          MoveL speed 75 mm/s, acceleration 150 mm/s^2 (useActiveTCP=true) feature=FRM_Reference
            SuppressedNode
              Script: PSE_T[2]=PSE_T[2]-0.005
            Waypoint Variable (Variable): variable=PSE_T
            SuppressedNode
              Force Frame feature=FRM_Reference; selection=[1, 1, 0, 0, 0, 0]; wrench=[0, 0, 0, 0, 0, 0]; limitsForce=[0.25, 0.25, 0.15, 1.047198, 1.047198, 1.047198]; limitsMotion=[0.1, 0.1, 0.1, 0.349066, 0.349066, 0.349066]
                Waypoint Variable (Variable): motionParameters(jointSpeed=1.047198 jointAcceleration=1.396263 cartesianSpeed=0.03 cartesianAcceleration=0.2); variable=PSE_T
            'ADD OPEN GRIPPER'
            Script: rq_set_force_norm(20)
            Script: rq_set_speed_norm(30)
            Script: rq_move_and_wait_norm(GRP_Close_Pos)
          Set DigitalOutput pin=digital_out[4]; digitalValue=1
          Wait Sleep waitTime=0.3
          MoveL speed 100 mm/s, acceleration 1200 mm/s^2 (useActiveTCP=true) feature=FRM_Reference
            Waypoint Variable (Variable): motionParameters(jointSpeed=1.047198 jointAcceleration=1.396263 cartesianSpeed=0.25 cartesianAcceleration=1.2); variable=PSE_R
      Case (caseValue=4)
        Folder Place probe in 3finger
          Action_Info := "place object"
          MoveJ speed 100 deg/s, acceleration 80 deg/s^2 (useActiveTCP=true) feature=FRM_Reference
            Waypoint Variable (Variable): variable=PSE_A
          Set DigitalOutput pin=digital_out[4]; digitalValue=1
          MoveL speed 75 mm/s, acceleration 150 mm/s^2 (useActiveTCP=true) feature=FRM_Reference
            Waypoint Variable (Variable): variable=PSE_T
              Until TOOL_CONTACT_DETECTION (allowActions=false retraction=0 decelerationAcceleration=3 decelerationAngularAcceleration=34.906585)
          Set DigitalOutput pin=digital_out[4]; digitalValue=0
          Wait Sleep waitTime=0.5
          SuppressedNode
            If Task_ID≟12
              Wait Sleep waitTime=0.15
              MoveL speed 75 mm/s, acceleration 150 mm/s^2 (useActiveTCP=true) feature=FRM_Reference
                Waypoint Variable (Variable): variable=PSE_R
      Case (caseValue=5)
        SuppressedNode
          Folder Decapping
            Action_Info := "decapping"
            PRM_decap_Zval := z_Pos
            PRM_forcdistSta := 0.02
            Script: zero_ftsensor()
            Wait Sleep waitTime=1
            Set DigitalOutput pin=digital_out[5]; digitalValue=1
            Set DigitalOutput pin=digital_out[3]; digitalValue=1
            Force Frame feature=uML_3fingergrip; selection=[0, 0, 1, 0, 0, 0]; wrench=[0, 0, 5, 0, 0, 0]; limitsForce=[0.04, 0.04, 0.015, 1.047198, 1.047198, 1.047198]; limitsMotion=[0.1, 0.1, 0.1, 0.349066, 0.349066, 0.349066]
              PRC_Force_Decap := True
              Wait Condition expression=PRM_forcdistLiv>PRM_forcdistSta
            PRC_Force_Decap := False
            Set DigitalOutput pin=digital_out[5]; digitalValue=0
            Set DigitalOutput pin=digital_out[3]; digitalValue=0
            MoveL speed 150 mm/s, acceleration 800 mm/s^2 (useActiveTCP=true) feature=FRM_Reference
              Waypoint Variable (Variable): variable=PSE_R
        Folder Decapping
          Action_Info := "decapping"
          Set DigitalOutput pin=digital_out[5]; digitalValue=1
          Set DigitalOutput pin=digital_out[3]; digitalValue=1
          Script: action_manipulator_decapping()
          Set DigitalOutput pin=digital_out[5]; digitalValue=0
          Set DigitalOutput pin=digital_out[3]; digitalValue=0
          MoveL speed 150 mm/s, acceleration 800 mm/s^2 (useActiveTCP=true) feature=FRM_Reference
            Waypoint Variable (Variable): variable=PSE_R
      Case (caseValue=6)
        SuppressedNode
          Folder Drop the cap
            Script: rq_set_speed_norm(100)
            Script: rq_set_force_norm(10)
            MoveJ speed 100 deg/s, acceleration 80 deg/s^2 (useActiveTCP=true) feature=FRM_Reference
              Waypoint Variable (Variable): motionParameters(blendRadius=0.02); variable=PSE_A
            MoveL speed 400 mm/s, acceleration 500 mm/s^2 (useActiveTCP=true) feature=FRM_Reference
              Waypoint Variable (Variable): motionParameters(jointSpeed=1.047198 jointAcceleration=1.396263 cartesianSpeed=0.09 cartesianAcceleration=0.05); variable=PSE_T
              'ADD OPEN GRIPPER'
              Loop While (checkContinuously=false) expression=rq_is_object_detected()
                URCap Gripper (Robotiq_Grippers, Robotiq Inc.) dataModel(position=0.0, force=28.0, speed=100.0, positionInDouble=0.0, forceInDouble=28.0, speedInDouble=100.0, slaveIds=[9], blocking=true)
                Wait Sleep waitTime=0.01
                URCap Gripper (Robotiq_Grippers, Robotiq Inc.) dataModel(position=100.0, force=28.0, speed=100.0, positionInDouble=100.0, forceInDouble=28.0, speedInDouble=100.0, slaveIds=[9], blocking=true)
              Wait Sleep waitTime=0.2
              Waypoint Variable (Variable): variable=PSE_R
        Folder Drop
          Script: rq_set_speed_norm(100)
          MoveJ speed 100 deg/s, acceleration 80 deg/s^2 (useActiveTCP=true) feature=FRM_Reference
            Waypoint Variable (Variable): motionParameters(blendRadius=0.02); variable=PSE_A
          MoveL speed 400 mm/s, acceleration 500 mm/s^2 (useActiveTCP=true) feature=FRM_Reference
            Waypoint Variable (Variable): motionParameters(jointSpeed=1.047198 jointAcceleration=1.396263 cartesianSpeed=0.12 cartesianAcceleration=0.08); variable=PSE_T
            URCap Gripper (Robotiq_Grippers, Robotiq Inc.) dataModel(position=70.19607843137254, force=30.19607843137255, speed=0.0, positionInDouble=70.19607843137254, forceInDouble=30.19607843137255, speedInDouble=0.0, slaveIds=[9], blocking=true)
            Waypoint Variable (Variable): motionParameters(jointSpeed=1.047198 jointAcceleration=1.396263 cartesianSpeed=0.12 cartesianAcceleration=0.08); variable=PSE_T_H
            Script: rq_move_and_wait_norm(GRP_Open_Pos)
            Wait Sleep waitTime=0.2
            Waypoint Variable (Variable): variable=PSE_R
      Case (caseValue=7)
        Folder Load
          Action_Info := "load object in the machine"
          SuppressedNode
            Script: do_transition(keep_rxry=OBJ_Picked)
          If JNT_Q≠JNT_Z
            Script: movej(get_inverse_kin(pose_trans(FRM_Reference, PSE_A), qnear=JNT_Q), r=0.05)
          Else 
            MoveJ speed 100 deg/s, acceleration 80 deg/s^2 (useActiveTCP=true) feature=FRM_Reference
              Waypoint Variable (Variable): motionParameters(blendRadius=0.02); variable=PSE_A
          MoveL speed 400 mm/s, acceleration 500 mm/s^2 (useActiveTCP=true) feature=FRM_Reference
            SuppressedNode
              Waypoint Variable (Variable): motionParameters(jointSpeed=1.047198 jointAcceleration=1.396263 cartesianSpeed=0.09 cartesianAcceleration=0.05); variable=PSE_T
                Until TOOL_CONTACT_DETECTION (allowActions=false retraction=0 decelerationAcceleration=0.5 decelerationAngularAcceleration=34.906585)
            SuppressedNode
              Force Frame feature=FRM_Reference; selection=[1, 1, 0, 0, 0, 0]; wrench=[0, 0, 0, 0, 0, 0]; limitsForce=[0.05, 0.05, 0.15, 1.047198, 1.047198, 1.047198]; limitsMotion=[0.1, 0.1, 0.1, 0.349066, 0.349066, 0.349066]
                Waypoint Variable (Variable): motionParameters(jointSpeed=1.047198 jointAcceleration=1.396263 cartesianSpeed=0.07 cartesianAcceleration=0.04); variable=PSE_T
            Waypoint Variable (Variable): motionParameters(jointSpeed=1.047198 jointAcceleration=1.396263 cartesianSpeed=0.07 cartesianAcceleration=0.04); variable=PSE_T_H
            URCap Gripper (Robotiq_Grippers, Robotiq Inc.) dataModel(position=100.0, force=0.0, speed=67.84313725490196, positionInDouble=100.0, forceInDouble=0.0, speedInDouble=67.84313725490196, slaveIds=[9], blocking=true)
            Wait Sleep waitTime=0.2
            Waypoint Variable (Variable): motionParameters(jointSpeed=1.047198 jointAcceleration=1.396263 cartesianSpeed=0.07 cartesianAcceleration=0.04); variable=PSE_T
            Waypoint Variable (Variable): variable=PSE_R
      Case (caseValue=8)
        Folder UnLoad
          Action_Info := "unload object in the machine"
          SuppressedNode
            Script: do_transition(keep_rxry=OBJ_Picked)
          If JNT_Q≠JNT_Z
            SuppressedNode
              Script: movej(get_inverse_kin(pose_trans(FRM_Reference, PSE_A), qnear=JNT_Q), r=0.01)
            Script: movej(get_inverse_kin(pose_trans(FRM_Reference, PSE_A), qnear=JNT_Q))
          Else 
            MoveJ speed 100 deg/s, acceleration 80 deg/s^2 (useActiveTCP=true) feature=FRM_Reference
              Waypoint Variable (Variable): variable=PSE_A
          MoveL speed 400 mm/s, acceleration 500 mm/s^2 (useActiveTCP=true) feature=FRM_Reference
            SuppressedNode
              Waypoint Variable (Variable): motionParameters(jointSpeed=1.047198 jointAcceleration=1.396263 cartesianSpeed=0.09 cartesianAcceleration=0.05); variable=PSE_T
                Until TOOL_CONTACT_DETECTION (allowActions=false retraction=0 decelerationAcceleration=0.5 decelerationAngularAcceleration=34.906585)
            SuppressedNode
              Force Frame feature=FRM_Reference; selection=[1, 1, 0, 0, 0, 0]; wrench=[0, 0, 0, 0, 0, 0]; limitsForce=[0.05, 0.05, 0.15, 1.047198, 1.047198, 1.047198]; limitsMotion=[0.1, 0.1, 0.1, 0.349066, 0.349066, 0.349066]
                Waypoint Variable (Variable): motionParameters(jointSpeed=1.047198 jointAcceleration=1.396263 cartesianSpeed=0.07 cartesianAcceleration=0.04); variable=PSE_T
            Script: rq_move_and_wait_norm(GRP_Open_Pos)
            Waypoint Variable (Variable): motionParameters(jointSpeed=1.047198 jointAcceleration=1.396263 cartesianSpeed=0.07 cartesianAcceleration=0.04); variable=PSE_T_H
            URCap Gripper (Robotiq_Grippers, Robotiq Inc.) dataModel(position=100.0, force=0.0, speed=67.84313725490196, positionInDouble=100.0, forceInDouble=0.0, speedInDouble=67.84313725490196, slaveIds=[9], blocking=true)
            Wait Sleep waitTime=0.2
            OBJ_Picked := rq_is_object_detected()
            If OBJ_Picked
              Waypoint Variable (Variable): motionParameters(jointSpeed=1.047198 jointAcceleration=1.396263 cartesianSpeed=0.07 cartesianAcceleration=0.04); variable=PSE_T
              Script: rq_move_and_wait_norm(GRP_Open_Pos)
              Waypoint Variable (Variable): variable=PSE_R
            Else 
              Script: set_error(1010)
      Case (caseValue=16)
        Folder Scan the barcode
          Action_Info := "scan the barcode"
          Barc_scan_succs := False
          Folder First check
            Set DigitalOutput pin=digital_out[6]; digitalValue=1
            Wait Sleep waitTime=0.1
            Barc_scan_succs := digital_in[6]
          If Barc_scan_succs
            Set DigitalOutput pin=digital_out[5]; digitalValue=1
            Set DigitalOutput pin=digital_out[2]; digitalValue=1
            Loop While (checkContinuously=true) expression=Barc_scan_succs
              Barc_scan_succs := digital_in[6]
              Wait Sleep waitTime=0.05
            Set DigitalOutput pin=digital_out[5]; digitalValue=0
            Set DigitalOutput pin=digital_out[2]; digitalValue=0
            Set DigitalOutput pin=digital_out[6]; digitalValue=0
          Else 
            Timer (action=Reset) variable=Timer_Barc_scan
            Timer (action=Start) variable=Timer_Barc_scan
            Set DigitalOutput pin=digital_out[3]; digitalValue=1
            Set DigitalOutput pin=digital_out[5]; digitalValue=1
            Loop While (checkContinuously=true) expression=not Barc_scan_succs and  not CMD_Stop and Timer_Barc_scan<60
              SuppressedNode
                If Timer_Barc_scan>1.5
                  Placeholder
              Set DigitalOutput pin=digital_out[6]; digitalValue=1
              Barc_scan_succs := digital_in[6]
              Wait Sleep waitTime=0.05
            Set DigitalOutput pin=digital_out[5]; digitalValue=0
            Set DigitalOutput pin=digital_out[3]; digitalValue=0
            Set DigitalOutput pin=digital_out[6]; digitalValue=0
            Timer (action=Stop) variable=Timer_Barc_scan
            If Timer_Barc_scan≥60
              Script: set_error(5200)
    '=========='
    Script: textmsg("Action=",Action)
    Folder PostSettings [hidden by the author, left out]
SubProgram Sub_AMR_MiR_V3 [hidden by the author, left out]
SubProgram Sub_Action_V4 (keepSynchronizedWithDisk=true) programFile=/programs/03 Sub Routines/Sub_Action_V4.urp
  Folder PreSettings
    Folder init poses [hidden by the author, left out]
    Folder Gripping parameters
      Script: OBJ = find_object_by_type(OBJs, OBJ_Type)
      GRP_Open_Pos := OBJ.dimension.diameter * 1000 + 6
      GRP_Offset := OBJ.gripper_offset
      Script: rq_set_force_norm(50)
      Script: rq_set_speed_norm(50)
    Switch expression=ITM_ID
      Case (caseValue=1)
        Folder uML
          Script: JIG2 = find_object_by_type(JIGs, JIG)
          JIG_Offset := JIG2.jig_offset
          Switch expression=JIG
            Case (caseValue=1)
              Folder 3FG
                Folder define poses
                  FRM_Reference := ULM_3FG
                  JNT_Q := JNT_HOME
                  PSE_T := pose_trans(GRP_Offset, JIG_Offset)
                  PSE_A := pose_trans(PSE_T, p[0,0,0.100,0,0,0])
                  PSE_R := pose_add(PSE_T, p[0,0,0.100,0,0,0])
            Case (caseValue=2)
              Folder Input
                'CHANGE THE REFERENCE TO THE FRAME TO MOVE IN'
                Folder define poses
                  FRM_Reference := ULM_Input
                  PSE_T := pose_trans(pose_trans(get_pattern_pos_rectangle(OBJ_Nbr, "X", [10,5], patternsize=[0.181,0.081]), GRP_Offset), JIG_Offset)
                  If Action≟1
                    PSE_R := pose_add(PSE_T, p[0,0,0.200,0,0,0])
                    PSE_A := pose_add(PSE_T, p[0,0,0.100,0,0,0])
                  ElseIf Action≟2
                    PSE_R := pose_add(PSE_T, p[0,0,0.100,0,0,0])
                    PSE_A := pose_add(PSE_T, p[0,0,0.200,0,0,0])
            Case (caseValue=3)
              Folder Output
                'CHANGE THE REFERENCE TO THE FRAME TO MOVE IN'
                Folder define poses
                  FRM_Reference := ULM_Output
                  PSE_T := pose_trans(pose_trans(get_pattern_pos_rectangle(OBJ_Nbr, "X", [10,5], patternsize=[0.181,0.081]), GRP_Offset), JIG_Offset)
                  SuppressedNode
                    PSE_T_H := 
                  If Action≟1
                    PSE_R := pose_add(PSE_T, p[0,0,0.200,0,0,0])
                    PSE_A := pose_add(PSE_T, p[0,0,0.100,0,0,0])
                  ElseIf Action≟2
                    PSE_R := pose_add(PSE_T, p[0,0,0.100,0,0,0])
                    PSE_A := pose_add(PSE_T, p[0,0,0.200,0,0,0])
            Case (caseValue=4)
              Folder jig centrifuge racks
                Folder define poses
                  FRM_Reference := ULM_Cent_Racks
                  PSE_T := get_pattern_pos_rectangle(JIG_Slot, "X", [4,1], patternsize=[0.291,0])
                  If OBJ_Nbr≠0
                    PSE_T := pose_trans(pose_trans(PSE_T, get_pattern_pos_rectangle(OBJ_Nbr, "X", [3,3], patternsize=[0.060,0.060])),p[-0.030, -0.030,0,0,0,3.927])
                  PSE_T := pose_trans(PSE_T, GRP_Offset)
                  If Action≟1
                    PSE_R := pose_add(PSE_T, p[0,0,0.200,0,0,0])
                    PSE_A := pose_add(PSE_T, p[0,0,0.100,0,0,0])
                  ElseIf Action≟2
                    PSE_R := pose_add(PSE_T, p[0,0,0.100,0,0,0])
                    PSE_A := pose_add(PSE_T, p[0,0,0.200,0,0,0])
            Case (caseValue=6)
              Folder Caps bin
                Folder define poses
                  'Drop cap'
                  Script: FRM_Reference=ULM_Cap_Bin
                  PSE_T := pose_RPY2RotVec(p[0,0,0,0,0,0])
                  PSE_T_H := pose_add(PSE_T, p[0,0,-0.011,0,0,0])
                  PSE_A := pose_trans(PSE_T, p[0,0,0.1,0,0,0])
                  PSE_R := pose_add(PSE_T, p[0,0,0.100,0,0,0])
            Case (caseValue=7)
              Folder Sarstedt
                'CHANGE THE REFERENCE TO THE FRAME TO MOVE IN'
                SuppressedNode
                  Folder Gripping parameters
                    GRP_Open_Pos := 45
                    GRP_Close_Pos := 100
                    Script: rq_set_force_norm(80)
                    Script: rq_set_speed_norm(100)
                If TASK.ID≟10
                  Folder Frame & Position Params
                    Script: FRM_Reference = ULM_SS_Rack
                    SuppressedNode
                      MoveL speed 250 mm/s, acceleration 1200 mm/s^2 (useActiveTCP=true) feature=FRM_Reference
                        Waypoint Variable (Variable): variable(featureName=uLM_SS_PickPlc)
                    SuppressedNode
                      PSE_T := pose_RPY2RotVec(p[0,0,0,0,0,0])
                    SuppressedNode
                      PSE_T := pose_trans(PSE_T, GRP_Offset)
                    PSE_T := uLM_SS_PickPlc
                    PSE_A := pose_trans(PSE_T, p[0,0,0.1,0,0,0])
                    PSE_R := pose_add(PSE_T, p[0,0,0.1,0,0,0])
                ElseIf TASK.ID≟11
                  Script: FRM_Reference = uLM_SS_PickPlc
                  PSE_T := pose_RPY2RotVec(p[0,0,0,0,0,0])
                  PSE_T := pose_trans(PSE_T, GRP_Offset)
                  PSE_A := pose_trans(PSE_T, p[0,0,0.1,0,0,0])
                  PSE_R := pose_add(PSE_T, p[0,0,0.2,0,0,0])
      Case (caseValue=2)
        Folder Centrifuge
          'CHANGE THE REFERENCE TO THE FRAME TO MOVE IN'
          Folder define poses
            FRM_Reference := FRM_Centrifuge
            PSE_T := GRP_Offset
            If Action≟8
              PSE_R := pose_add(PSE_T, p[0,0,0.250,0,0,0])
              PSE_A := pose_add(PSE_T, p[0,0,0.150,0,0,0])
            ElseIf Action≟7
              PSE_R := pose_add(PSE_T, p[0,0,0.150,0,0,0])
              PSE_A := pose_add(PSE_T, p[0,0,0.250,0,0,0])
      Case (caseValue=3)
        Folder Output
          'CHANGE THE REFERENCE TO THE FRAME TO MOVE IN'
          Folder define poses
            FRM_Reference := Base
            PSE_T := p[0,0,0,0,0,0]
            PSE_A := pose_add(PSE_T, p[0,0,0.150,0,0,0])
            PSE_R := pose_add(PSE_T, p[0,0,0.100,0,0,0])
      Case (caseValue=5)
        Folder Sarstedt Pickup Table
          'CHANGE THE REFERENCE TO THE FRAME TO MOVE IN'
          Switch expression=JIG
            Case (caseValue=7)
              Folder Sarstedt Rack
                SuppressedNode
                  Folder Gripping parameters
                    GRP_Open_Pos := 45
                    GRP_Close_Pos := 100
                    Script: rq_set_force_norm(80)
                    Script: rq_set_speed_norm(100)
                Folder Frame & Position Params
                  Script: FRM_Reference = FRM_SS_SSTable
                  PSE_T := pose_RPY2RotVec(p[0,0,0,0,0,0])
                  PSE_T := pose_trans(PSE_T, GRP_Offset)
                  PSE_A := pose_trans(PSE_T, p[0,0,0.1,0,0,0])
                  PSE_R := pose_add(PSE_T, p[0,0,0.1,0,0,0])
    Folder Additional check [hidden by the author, left out]
  '=========='
  Switch expression=Action
    Case (caseValue=1)
      Folder Pick
        Action_Info := "pick object"
        Script: do_transition(pose_trans(FRM_Reference, PSE_T), keep_rxry=OBJ_Picked)
        Folder EOAT
          If not OBJ_Picked
            Script: rq_move_and_wait_mm(GRP_Open_Pos)
        If PSE_A_H≠PSE_Z
          If JNT_Q≠JNT_Z
            Script: movej(get_inverse_kin(pose_trans(FRM_Reference, PSE_A_H), qnear=JNT_Q), r=0.050)
          Else 
            Script: movej(pose_trans(FRM_Reference, PSE_A_H), r=0.050)
        If PSE_A≠PSE_Z
          If JNT_Q≠JNT_Z
            Script: movej(get_inverse_kin(pose_trans(FRM_Reference, PSE_A), qnear=JNT_Q), r=0.020)
          Else 
            Script: movej(pose_trans(FRM_Reference, PSE_A), r=0.020)
        MoveL speed 400 mm/s, acceleration 500 mm/s^2 (useActiveTCP=true) feature=FRM_Reference
          If PSE_T_H≠PSE_Z
            Waypoint Variable (Variable): motionParameters(blendRadius=0.01); variable=PSE_T_H
          Waypoint Variable (Variable): motionParameters(jointSpeed=1.047198 jointAcceleration=1.396263 cartesianSpeed=0.12 cartesianAcceleration=0.08); variable=PSE_T
          Folder EOAT
            Script: rq_set_force_norm(50)
            Script: rq_close_and_wait()
            OBJ_Picked := rq_is_object_detected()
            If not OBJ_Picked
              Script: set_error(ERROR_NO_OBJECT_TO_PICK)
          Folder EXTT
            Switch expression=JIG
              Case (caseValue=1)
                Folder 3FG
                  If OBJ_Picked
                    Set DigitalOutput pin=digital_out[5]; digitalValue=1
          If PSE_R_H≠PSE_Z
            Waypoint Variable (Variable): motionParameters(blendRadius=0.01); variable=PSE_R
            Waypoint Variable (Variable): variable=PSE_R_H
          Else 
            Waypoint Variable (Variable): variable=PSE_R
    Case (caseValue=2)
      Folder Place
        Action_Info := "place object"
        Script: do_transition(pose_trans(FRM_Reference, PSE_T), keep_rxry=OBJ_Picked)
        Folder EXTT
          Switch expression=JIG
            Case (caseValue=1)
              Folder 3FG
                If OBJ_Picked
                  Set DigitalOutput pin=digital_out[5]; digitalValue=1
        If PSE_A_H≠PSE_Z
          If JNT_Q≠JNT_Z
            Script: movej(get_inverse_kin(pose_trans(FRM_Reference, PSE_A_H), qnear=JNT_Q), r=0.050)
          Else 
            Script: movej(pose_trans(FRM_Reference, PSE_A_H), r=0.050)
        If PSE_A≠PSE_Z
          If JNT_Q≠JNT_Z
            Script: movej(get_inverse_kin(pose_trans(FRM_Reference, PSE_A), qnear=JNT_Q), r=0.020)
          Else 
            Script: movej(pose_trans(FRM_Reference, PSE_A), r=0.020)
        MoveL speed 400 mm/s, acceleration 500 mm/s^2 (useActiveTCP=true) feature=FRM_Reference
          If PSE_T_H≠PSE_Z
            Waypoint Variable (Variable): motionParameters(blendRadius=0.01); variable=PSE_T_H
          Waypoint Variable (Variable): motionParameters(jointSpeed=1.047198 jointAcceleration=1.396263 cartesianSpeed=0.09 cartesianAcceleration=0.05); variable=PSE_T
            Until TOOL_CONTACT_DETECTION (allowActions=false retraction=NONE decelerationAcceleration=0.5 decelerationAngularAcceleration=34.906585)
          Force Frame feature=FRM_Reference; selection=[1, 1, 1, 0, 0, 0]; wrench=[0, 0, 0, 0, 0, 0]; limitsForce=[0.1, 0.1, 0.01, 1.047198, 1.047198, 1.047198]; limitsMotion=[0.1, 0.1, 0.1, 0.349066, 0.349066, 0.349066]
            Waypoint Variable (Variable): motionParameters(jointSpeed=1.047198 jointAcceleration=1.396263 cartesianSpeed=0.07 cartesianAcceleration=0.04); variable=PSE_T
          Folder EXTT
            Switch expression=JIG
              Case (caseValue=1)
                Folder 3FG
                  If OBJ_Picked
                    Set DigitalOutput pin=digital_out[5]; digitalValue=0
                    Wait Sleep waitTime=0.2
          Folder EOAT
            Script: rq_move_and_wait_mm(GRP_Open_Pos)
            OBJ_Picked := rq_is_object_detected()
          If PSE_R_H≠PSE_Z
            Waypoint Variable (Variable): motionParameters(blendRadius=0.01); variable=PSE_R
            Waypoint Variable (Variable): variable=PSE_R_H
          Else 
            Waypoint Variable (Variable): variable=PSE_R
    Case (caseValue=3)
      Folder Push
        Action_Info := "push"
    Case (caseValue=4)
      Folder Pull
        Action_Info := "pull"
    SuppressedNode
      Case (caseValue=5)
        Placeholder
    Case (caseValue=6)
      SuppressedNode
        Folder Drop the cap
          If JNT_A≠[0,0,0,0,0,0]
            MoveJ speed 100 deg/s, acceleration 80 deg/s^2 (useActiveTCP=true positionType=JointAngles) feature=FRM_Reference
              Waypoint Variable (Variable): motionParameters(blendRadius=0.02); variable=JNT_A
          Else 
            MoveJ speed 100 deg/s, acceleration 80 deg/s^2 (useActiveTCP=true) feature=FRM_Reference
              Waypoint Variable (Variable): motionParameters(blendRadius=0.02); variable=PSE_A
          MoveL speed 400 mm/s, acceleration 500 mm/s^2 (useActiveTCP=true) feature=FRM_Reference
            Waypoint Variable (Variable): motionParameters(jointSpeed=1.047198 jointAcceleration=1.396263 cartesianSpeed=0.09 cartesianAcceleration=0.05); variable=PSE_T
            'ADD OPEN GRIPPER'
            URCap Gripper (Robotiq_Grippers, Robotiq Inc.) dataModel(position=78.82352941176471, force=11.0, speed=0.0, positionInDouble=78.82352941176471, forceInDouble=11.0, speedInDouble=0.0, slaveIds=[9], blocking=true)
            Waypoint Variable (Variable): motionParameters(jointSpeed=1.047198 jointAcceleration=1.396263 cartesianSpeed=0.09 cartesianAcceleration=0.05); variable=PSE_T_H
            URCap Gripper (Robotiq_Grippers, Robotiq Inc.) dataModel(position=24.705882352941178, force=11.0, speed=0.0, positionInDouble=24.705882352941178, forceInDouble=11.0, speedInDouble=0.0, slaveIds=[9], blocking=true)
            SuppressedNode
              URCap Gripper (Robotiq_Grippers, Robotiq Inc.) dataModel(position=100.0, force=28.0, speed=100.0, positionInDouble=100.0, forceInDouble=28.0, speedInDouble=100.0, slaveIds=[9], blocking=true)
            SuppressedNode
              Wait Sleep waitTime=0.2
            SuppressedNode
              Loop While (checkContinuously=false) expression=rq_is_object_detected()
                Script: rq_set_force_norm(10)
                Script: rq_set_speed_norm(100)
                URCap Gripper (Robotiq_Grippers, Robotiq Inc.) dataModel(position=0.0, force=28.0, speed=100.0, positionInDouble=0.0, forceInDouble=28.0, speedInDouble=100.0, slaveIds=[9], blocking=true)
                Wait Sleep waitTime=0.5
                URCap Gripper (Robotiq_Grippers, Robotiq Inc.) dataModel(position=100.0, force=28.0, speed=100.0, positionInDouble=100.0, forceInDouble=28.0, speedInDouble=100.0, slaveIds=[9], blocking=true)
            SuppressedNode
              Wait Sleep waitTime=0.2
            Waypoint Variable (Variable): variable=PSE_R
    Case (caseValue=7)
      Folder Load
        Action_Info := "load object"
        Script: do_transition(pose_trans(FRM_Reference, PSE_T), keep_rxry=OBJ_Picked)
        If PSE_A_H≠PSE_Z
          If JNT_Q≠JNT_Z
            Script: movej(get_inverse_kin(pose_trans(FRM_Reference, PSE_A_H), qnear=JNT_Q), r=0.050)
          Else 
            Script: movej(pose_trans(FRM_Reference, PSE_A_H), r=0.050)
        If PSE_A≠PSE_Z
          If JNT_Q≠JNT_Z
            Script: movej(get_inverse_kin(pose_trans(FRM_Reference, PSE_A), qnear=JNT_Q), r=0.020)
          Else 
            Script: movej(pose_trans(FRM_Reference, PSE_A), r=0.020)
        MoveL speed 400 mm/s, acceleration 500 mm/s^2 (useActiveTCP=true) feature=FRM_Reference
          If PSE_T_H≠PSE_Z
            Waypoint Variable (Variable): motionParameters(blendRadius=0.01); variable=PSE_T_H
          Waypoint Variable (Variable): motionParameters(jointSpeed=1.047198 jointAcceleration=1.396263 cartesianSpeed=0.09 cartesianAcceleration=0.05); variable=PSE_T
            Until TOOL_CONTACT_DETECTION (allowActions=false retraction=NONE decelerationAcceleration=0.5 decelerationAngularAcceleration=34.906585)
          Force Frame feature=FRM_Reference; selection=[0, 1, 1, 0, 0, 1]; wrench=[0, 0, 0, 0, 0, 0]; limitsForce=[0.1, 0.05, 0.02, 1.047198, 1.047198, 3.141593]; limitsMotion=[0.1, 0.1, 0.1, 0.349066, 0.349066, 0.349066]
            Waypoint Variable (Variable): motionParameters(jointSpeed=1.047198 jointAcceleration=1.396263 cartesianSpeed=0.07 cartesianAcceleration=0.04); variable=PSE_T
          Folder EOAT
            Script: rq_move_and_wait_mm(GRP_Open_Pos)
            OBJ_Picked := rq_is_object_detected()
          If PSE_R_H≠PSE_Z
            Waypoint Variable (Variable): motionParameters(blendRadius=0.01); variable=PSE_R
            Waypoint Variable (Variable): variable=PSE_R_H
          Else 
            Waypoint Variable (Variable): variable=PSE_R
    Case (caseValue=8)
      Folder Unload
        Action_Info := "pick object"
        Script: do_transition(pose_trans(FRM_Reference, PSE_T), keep_rxry=OBJ_Picked)
        Folder EOAT
          If not OBJ_Picked
            Script: rq_move_and_wait_mm(GRP_Open_Pos)
        If PSE_A_H≠PSE_Z
          If JNT_Q≠JNT_Z
            Script: movej(get_inverse_kin(pose_trans(FRM_Reference, PSE_A_H), qnear=JNT_Q), r=0.050)
          Else 
            Script: movej(pose_trans(FRM_Reference, PSE_A_H), r=0.050)
        If PSE_A≠PSE_Z
          If JNT_Q≠JNT_Z
            Script: movej(get_inverse_kin(pose_trans(FRM_Reference, PSE_A), qnear=JNT_Q), r=0.020)
          Else 
            Script: movej(pose_trans(FRM_Reference, PSE_A), r=0.020)
        MoveL speed 400 mm/s, acceleration 500 mm/s^2 (useActiveTCP=true) feature=FRM_Reference
          If PSE_T_H≠PSE_Z
            Waypoint Variable (Variable): motionParameters(blendRadius=0.01); variable=PSE_T_H
          Waypoint Variable (Variable): motionParameters(jointSpeed=1.047198 jointAcceleration=1.396263 cartesianSpeed=0.12 cartesianAcceleration=0.08); variable=PSE_T
          Force Frame feature=FRM_Reference; selection=[1, 1, 0, 0, 0, 0]; wrench=[0, 0, 0, 0, 0, 0]; limitsForce=[0.05, 0.05, 0.15, 1.047198, 1.047198, 1.047198]; limitsMotion=[0.1, 0.1, 0.1, 0.349066, 0.349066, 0.349066]
            Folder EOAT
              Script: rq_set_force_norm(50)
              Script: rq_close_and_wait()
              OBJ_Picked := rq_is_object_detected()
              If not OBJ_Picked
                Script: set_error(ERROR_NO_OBJECT_TO_PICK)
            If PSE_R_H≠PSE_Z
              Waypoint Variable (Variable): motionParameters(blendRadius=0.01); variable=PSE_R
              Waypoint Variable (Variable): variable=PSE_R_H
            Else 
              Waypoint Variable (Variable): variable=PSE_R
    Case (caseValue=11)
      Folder Place
        Action_Info := "place object without gripper opening"
        Script: do_transition(pose_trans(FRM_Reference, PSE_T), keep_rxry=OBJ_Picked)
        Folder EXTT
          Switch expression=JIG
            Case (caseValue=1)
              Folder 3FG
                If OBJ_Picked
                  Set DigitalOutput pin=digital_out[5]; digitalValue=1
        If PSE_A_H≠PSE_Z
          If JNT_Q≠JNT_Z
            Script: movej(get_inverse_kin(pose_trans(FRM_Reference, PSE_A_H), qnear=JNT_Q), r=0.050)
          Else 
            Script: movej(pose_trans(FRM_Reference, PSE_A_H), r=0.050)
        If PSE_A≠PSE_Z
          If JNT_Q≠JNT_Z
            Script: movej(get_inverse_kin(pose_trans(FRM_Reference, PSE_A), qnear=JNT_Q), r=0.020)
          Else 
            Script: movej(pose_trans(FRM_Reference, PSE_A), r=0.020)
        MoveL speed 400 mm/s, acceleration 500 mm/s^2 (useActiveTCP=true) feature=FRM_Reference
          If PSE_T_H≠PSE_Z
            Waypoint Variable (Variable): motionParameters(blendRadius=0.01); variable=PSE_T_H
          Waypoint Variable (Variable): motionParameters(jointSpeed=1.047198 jointAcceleration=1.396263 cartesianSpeed=0.09 cartesianAcceleration=0.05); variable=PSE_T
            Until TOOL_CONTACT_DETECTION (allowActions=false retraction=NONE decelerationAcceleration=0.5 decelerationAngularAcceleration=34.906585)
          Force Frame feature=FRM_Reference; selection=[1, 1, 1, 0, 0, 0]; wrench=[0, 0, 0, 0, 0, 0]; limitsForce=[0.1, 0.1, 0.01, 1.047198, 1.047198, 1.047198]; limitsMotion=[0.1, 0.1, 0.1, 0.349066, 0.349066, 0.349066]
            Waypoint Variable (Variable): motionParameters(jointSpeed=1.047198 jointAcceleration=1.396263 cartesianSpeed=0.07 cartesianAcceleration=0.04); variable=PSE_T
          Folder EXTT
            Switch expression=JIG
              Case (caseValue=1)
                Folder 3FG
                  If OBJ_Picked
                    Set DigitalOutput pin=digital_out[5]; digitalValue=0
                    Wait Sleep waitTime=0.2
          Folder EOAT
            ''
    Case (caseValue=12)
      Folder Decap
        Action_Info := "decapping"
        Set DigitalOutput pin=digital_out[4]; digitalValue=1
        Set DigitalOutput pin=digital_out[3]; digitalValue=1
        Force Simple feature=Joint_6_name; selection=[0, 0, 1, 0, 0, 0]; wrench=[0, 0, 5, 0, 0, 0]; limitsForce=[0.15, 0.15, 0.15, 1.047198, 1.047198, 1.047198]; limitsMotion=[0.1, 0.1, 0.1, 0.349066, 0.349066, 0.349066]
          Script: check_decapping(offset=0.015, timeout=5, abort=CMD_Hold)
        Set DigitalOutput pin=digital_out[3]; digitalValue=0
        Set DigitalOutput pin=digital_out[4]; digitalValue=0
        MoveL speed 150 mm/s, acceleration 800 mm/s^2 (useActiveTCP=true) feature=FRM_Reference
          Waypoint Variable (Variable): variable=PSE_R
    Case (caseValue=13)
      SuppressedNode
        Folder Read
          Folder Search for code
            Wait Condition expression=( not digital_in[6] and  not Barcode_nOK and  not digital_out[3])
            Timer (action=Start) variable(name=TMR_Barcode)
            Set DigitalOutput pin=digital_out[2]; digitalValue=1
            Set DigitalOutput pin=digital_out[6]; digitalValue=1
            Wait Condition expression=TMR_Barcode≥PRM_TO_Read_BC or digital_in[6] or Barcode_nOK
            Set DigitalOutput pin=digital_out[2]; digitalValue=0
            Set DigitalOutput pin=digital_out[6]; digitalValue=0
            Timer (action=Stop) variable=TMR_Barcode
          If digital_in[6]
            Folder barcode found
              'nothing'
          ElseIf Barcode_nOK or TMR_Barcode≥PRM_TO_Read_BC
            Placeholder
      Timer (action=Reset) variable=TMR_Barcode
      Folder Read
        Timer (action=Start) variable=TMR_Barcode
        If TMR_Barcode<PRM_TO_Read_BC
          Folder KeyenceTrigger
            Set SingleDigitalPulseActionState SingleDigitalPulseActionState(hiPulseInSeconds=0.2, pin=GP_bool_out[2])
            Wait Sleep waitTime=0.5
            Set DigitalOutput pin=GP_bool_out[1]; digitalValue=0
            Wait Sleep waitTime=0.5
            Set DigitalOutput pin=GP_bool_out[1]; digitalValue=1
            Wait Sleep waitTime=0.5
          Folder Preorient
            Timer (action=Reset) variable=TMR_Barcode
            If GP_bool_in[12]
              Set DigitalOutput pin=digital_out[3]; digitalValue=1
              Set DigitalOutput pin=digital_out[4]; digitalValue=1
              Loop While (checkContinuously=false) expression=GP_bool_in[12]
                Folder KeyenceTrigger
                  Set SingleDigitalPulseActionState SingleDigitalPulseActionState(hiPulseInSeconds=0.1, pin=GP_bool_out[2])
                  Wait Sleep waitTime=0.3
                  Set DigitalOutput pin=GP_bool_out[1]; digitalValue=0
                  Wait Sleep waitTime=0.3
                  Set DigitalOutput pin=GP_bool_out[1]; digitalValue=1
                  Wait Sleep waitTime=0.1
            If not GP_bool_in[12]
              Set DigitalOutput pin=digital_out[3]; digitalValue=1
              Set DigitalOutput pin=digital_out[4]; digitalValue=1
              Wait DigitalInput pin=GP_bool_in[12]; digitalValue=1
          Set DigitalOutput pin=digital_out[3]; digitalValue=0
          Set DigitalOutput pin=digital_out[4]; digitalValue=0
        Else 
          Folder exeption
            Folder error
              Script: set_error(6000)
        Set DigitalOutput pin=digital_out[3]; digitalValue=0
        Set DigitalOutput pin=digital_out[4]; digitalValue=0
        Set DigitalOutput pin=GP_bool_out[1]; digitalValue=0
    Case (caseValue=15)
      Folder Detect [hidden by the author, left out]
  '=========='
  Folder PostSettings [hidden by the author, left out]
